(*
SPDX-FileCopyrightText: c 2026 Oleksandr Tiutyk <trofimich@gmail.com>
SPDX-License-Identifier: MIT
License: https://opensource.org/license/mit
*)

(*!
<summary>Exercises all five native event categories.</summary>
<description>
Each run submits five numbered messages from the runner task and checks each admission result.
</description>
*)

{attribute 'no_assign'}
{attribute 'no_explicit_call' := 'do not call this function block directly'}
FUNCTION_BLOCK EventLoggerCategoryTest EXTENDS TOF_Testing.SingleCycleTest
VAR_STAT
	{attribute 'hide'}
	_ClassName : STRING := __POUNAME();
END_VAR
VAR
	_EventLogger : TOF_Loggers.EventLogger(
		debugEventType := TC_EVENTS.OpenFrameworkLoggerEventClass.DebugEvent,
		informationEventType := TC_EVENTS.OpenFrameworkLoggerEventClass.InformationEvent,
		warningEventType := TC_EVENTS.OpenFrameworkLoggerEventClass.WarningEvent,
		errorEventType := TC_EVENTS.OpenFrameworkLoggerEventClass.ErrorEvent,
		criticalErrorEventType := TC_EVENTS.OpenFrameworkLoggerEventClass.CriticalErrorEvent
	);
END_VAR

(*!
<summary>Sends a numbered message for each configured event type and checks the native result.</summary>
*)
METHOD PROTECTED ExecuteTest
VAR
	number : ULINT;
END_VAR
number := 1;
Assert.ThatBool(
	actual := _EventLogger.TryLogMessage(
		category := TOF_Core.LOG_CATEGORY.DEBUG,
		message := "LoggerTest DEBUG",
		messageNumber := number
	),
	message := "EventLogger refused DEBUG"
).IsTrue();

number := 2;
Assert.ThatBool(
	actual := _EventLogger.TryLogMessage(
		category := TOF_Core.LOG_CATEGORY.INFORMATION,
		message := "LoggerTest INFORMATION",
		messageNumber := number
	),
	message := "EventLogger refused INFORMATION"
).IsTrue();

number := 3;
Assert.ThatBool(
	actual := _EventLogger.TryLogMessage(
		category := TOF_Core.LOG_CATEGORY.WARNING,
		message := "LoggerTest WARNING",
		messageNumber := number
	),
	message := "EventLogger refused WARNING"
).IsTrue();

number := 4;
Assert.ThatBool(
	actual := _EventLogger.TryLogMessage(
		category := TOF_Core.LOG_CATEGORY.ERROR,
		message := "LoggerTest ERROR",
		messageNumber := number
	),
	message := "EventLogger refused ERROR"
).IsTrue();

number := 5;
Assert.ThatBool(
	actual := _EventLogger.TryLogMessage(
		category := TOF_Core.LOG_CATEGORY.CRITICAL_ERROR,
		message := "LoggerTest CRITICAL_ERROR",
		messageNumber := number
	),
	message := "EventLogger refused CRITICAL_ERROR"
).IsTrue();
END_METHOD

//! <summary>Borrows the concrete class name for the instance lifetime. Callers must not modify it.</summary>
{attribute 'monitoring' := 'call'}
PROPERTY ClassName : REFERENCE TO STRING
GET
ClassName REF= _ClassName;
END_GET
END_PROPERTY

//! <summary>Borrows the compiler-initialized namespace. Callers must not modify it.</summary>
{attribute 'monitoring' := 'call'}
PROPERTY NamespaceName : REFERENCE TO STRING
GET
NamespaceName REF= CurrentNamespace.Name;
END_GET
END_PROPERTY

//! <summary>Reports the complete instance size in bytes, excluding separately allocated storage.</summary>
{attribute 'monitoring' := 'call'}
PROPERTY SelfSize : ULINT
GET
SelfSize := XSIZEOF(THIS^);
END_GET
END_PROPERTY

END_FUNCTION_BLOCK

(* stored: Version 1.1.0.1
   POU EventLoggerCategoryTest: Id {a11e9240-740e-49fe-a8bc-709cb7f36a7c}, SpecialFunc None
   Method ExecuteTest: Id {049cb0f6-6383-4bca-a941-6faedabca72c}
   Property ClassName: Id {4d1a30ad-5cd6-4d2c-b459-12188e7a8e3f}
   Get Get: Id {98f6f448-a343-427d-8030-747d66cb901e}
   Property NamespaceName: Id {67b035d9-d1df-4178-953d-ecf32d34e0a2}
   Get Get: Id {7dd4cd35-4021-4f1d-9041-634f20b5a721}
   Property SelfSize: Id {3b7ec68f-30fb-411b-b0dd-70ef7cec62f0}
   Get Get: Id {327d1e76-eb0b-4422-b918-bbacdb001da8} *)
